TYPE ST_DeviceErrorHandeling :
STRUCT
	eName			: E_OwnerDevice:=E_OwnerDevice.NotDefined;
	sObjectName		: STRING:='Device Name';
	iObjectID		: INT;
	sLastErrorStep	: STRING;
	eErrorActive	: E_Error_Active_Module:=E_Error_Active_Module.noError;
	bMasterResume	: BOOL;

END_STRUCT
END_TYPE

(* stored: Version 1.1.0.1, ProductVersion 3.1.4024.12
   DUT ST_DeviceErrorHandeling: Id {552268b2-db52-4082-bb49-8cc4726470df} *)
